(* IEC 61131-3 sources: rusty/tests/lit/single/polymorphism/interfaces, 25 files *)

(* ---- argument.st ---- *)
// RUN: %COMPILE %s && %RUN | %CHECK %s
// Scenario: Ensure interface references passed as VAR_INPUT arguments are correctly dispatched to the
// implementing function block's method.

INTERFACE IA
    METHOD foo
    END_METHOD
END_INTERFACE

INTERFACE IB
    METHOD bar
        VAR_INPUT
            refIA: IA;
        END_VAR
    END_METHOD
END_INTERFACE

FUNCTION_BLOCK FbA IMPLEMENTS IA
    METHOD foo
        printf('FbA::foo$N');
    END_METHOD
END_FUNCTION_BLOCK

FUNCTION_BLOCK FbB IMPLEMENTS IB
    VAR_INPUT
        refIA: IA;
    END_VAR

    METHOD bar
        VAR_INPUT
            refIA: IA;
        END_VAR

        refIA.foo();
        printf('FbB::bar$N');
    END_METHOD

    refIA.foo();
END_FUNCTION_BLOCK

FUNCTION main
    VAR
        instanceFbA: FbA;
        instanceFbB: FbB;
    END_VAR

    // CHECK: FbA::foo
    instanceFbB(refIA := instanceFbA);

    // CHECK-NEXT: FbA::foo
    // CHECK-NEXT: FbB::bar
    instanceFbB.bar(refIA := instanceFbA);
END_FUNCTION

(* ---- argument_implicit.st ---- *)
// RUN: %COMPILE %s && %RUN | %CHECK %s
// Scenario: FbA implements IA, FbB extends FbA and implicitly implements IA. Both should be passable as
// interface-typed arguments, with FbB's overridden method dispatched correctly.

INTERFACE IA
    METHOD foo
    END_METHOD
END_INTERFACE

FUNCTION_BLOCK FbA IMPLEMENTS IA
    METHOD foo
        printf('FbA::foo$N');
    END_METHOD
END_FUNCTION_BLOCK

FUNCTION_BLOCK FbB EXTENDS FbA
    METHOD foo
        printf('FbB::foo$N');
    END_METHOD
END_FUNCTION_BLOCK

FUNCTION_BLOCK FbC EXTENDS FbB
END_FUNCTION_BLOCK

FUNCTION_BLOCK FbConsumer
    METHOD bar
        VAR_INPUT
            refIA: IA;
        END_VAR

        refIA.foo();
    END_METHOD
END_FUNCTION_BLOCK

FUNCTION main
    VAR
        instanceFbA: FbA;
        instanceFbB: FbB;
        instanceFbC: FbC;
        consumer: FbConsumer;
    END_VAR

    // CHECK: FbA::foo
    consumer.bar(refIA := instanceFbA);

    // CHECK-NEXT: FbB::foo
    consumer.bar(refIA := instanceFbB);

    // FbC inherits FbB's override
    // CHECK-NEXT: FbB::foo
    consumer.bar(refIA := instanceFbC);
END_FUNCTION

(* ---- argument_mixed.st ---- *)
// RUN: %COMPILE %s && %RUN | %CHECK %s
// Scenario: A method takes a mix of interface-typed and non-interface-typed parameters. Only the
// interface-typed arguments should be wrapped in a fat pointer; the rest remain untouched.

INTERFACE IA
    METHOD foo
    END_METHOD
END_INTERFACE

FUNCTION_BLOCK FbA IMPLEMENTS IA
    METHOD foo
        printf('FbA::foo$N');
    END_METHOD
END_FUNCTION_BLOCK

FUNCTION_BLOCK FbConsumer
    METHOD bar
        VAR_INPUT
            x: DINT;
            refIA: IA;
            y: DINT;
        END_VAR

        printf('x=%d, y=%d$N', x, y);
        refIA.foo();
    END_METHOD
END_FUNCTION_BLOCK

FUNCTION main
    VAR
        instanceFbA: FbA;
        consumer: FbConsumer;
    END_VAR

    // CHECK: x=1, y=2
    // CHECK-NEXT: FbA::foo
    consumer.bar(x := 1, refIA := instanceFbA, y := 2);
END_FUNCTION

(* ---- argument_positional.st ---- *)
// RUN: %COMPILE %s && %RUN | %CHECK %s
// Scenario: Interface references passed as positional (unnamed) VAR_INPUT arguments are correctly wrapped
// in a fat pointer and dispatched to the implementing function block's method.

INTERFACE IA
    METHOD foo
    END_METHOD
END_INTERFACE

FUNCTION_BLOCK FbA IMPLEMENTS IA
    METHOD foo
        printf('FbA::foo$N');
    END_METHOD
END_FUNCTION_BLOCK

FUNCTION_BLOCK FbB IMPLEMENTS IA
    METHOD foo
        printf('FbB::foo$N');
    END_METHOD
END_FUNCTION_BLOCK

FUNCTION_BLOCK FbConsumer
    METHOD bar
        VAR_INPUT
            refIA: IA;
        END_VAR

        refIA.foo();
    END_METHOD
END_FUNCTION_BLOCK

FUNCTION main
    VAR
        instanceFbA: FbA;
        instanceFbB: FbB;
        consumer: FbConsumer;
    END_VAR

    // CHECK: FbA::foo
    consumer.bar(instanceFbA);

    // CHECK-NEXT: FbB::foo
    consumer.bar(instanceFbB);
END_FUNCTION

(* ---- argument_sequential.st ---- *)
// RUN: %COMPILE %s && %RUN | %CHECK %s
// Scenario: Multiple sequential calls pass different concrete types to the same interface-typed parameter.
// The single __tmp variable is reused across calls — each call should dispatch to the correct implementation.

INTERFACE IA
    METHOD foo
    END_METHOD
END_INTERFACE

FUNCTION_BLOCK FbA IMPLEMENTS IA
    METHOD foo
        printf('FbA::foo$N');
    END_METHOD
END_FUNCTION_BLOCK

FUNCTION_BLOCK FbB IMPLEMENTS IA
    METHOD foo
        printf('FbB::foo$N');
    END_METHOD
END_FUNCTION_BLOCK

FUNCTION_BLOCK FbC IMPLEMENTS IA
    METHOD foo
        printf('FbC::foo$N');
    END_METHOD
END_FUNCTION_BLOCK

FUNCTION_BLOCK FbConsumer
    METHOD bar
        VAR_INPUT
            refIA: IA;
        END_VAR

        refIA.foo();
    END_METHOD
END_FUNCTION_BLOCK

FUNCTION main
    VAR
        instanceFbA: FbA;
        instanceFbB: FbB;
        instanceFbC: FbC;
        consumer: FbConsumer;
    END_VAR

    // CHECK: FbA::foo
    consumer.bar(refIA := instanceFbA);

    // CHECK-NEXT: FbB::foo
    consumer.bar(refIA := instanceFbB);

    // CHECK-NEXT: FbC::foo
    consumer.bar(refIA := instanceFbC);

    // Back to FbA to confirm __tmp is correctly overwritten
    // CHECK-NEXT: FbA::foo
    consumer.bar(refIA := instanceFbA);
END_FUNCTION

(* ---- combined_aggregate_return_mixed_args.st ---- *)
// RUN: %COMPILE %s && %RUN | %CHECK %s
// Scenario: A method returns a STRUCT (aggregate) and takes a mix of scalar, interface, and multiple
// different interface-typed parameters. Tests both positional (unnamed) and named arguments with
// completely reordered parameter positions to verify that fat pointer wrapping targets the correct
// parameters regardless of call-site argument order.

TYPE Result :
    STRUCT
        summary: STRING;
        total: DINT;
    END_STRUCT
END_TYPE

INTERFACE IA
    METHOD describe : STRING
    END_METHOD
END_INTERFACE

INTERFACE IB
    METHOD value : DINT
    END_METHOD
END_INTERFACE

INTERFACE IC
    METHOD combine : Result
        VAR_INPUT
            x: DINT;
            a: IA;
            y: REAL;
            b: IB;
            label: STRING;
        END_VAR
    END_METHOD
END_INTERFACE

FUNCTION_BLOCK FbA IMPLEMENTS IA
    METHOD describe : STRING
        describe := 'FbA';
    END_METHOD
END_FUNCTION_BLOCK

FUNCTION_BLOCK FbB IMPLEMENTS IB
    METHOD value : DINT
        value := 100;
    END_METHOD
END_FUNCTION_BLOCK

FUNCTION_BLOCK FbC IMPLEMENTS IC
    METHOD combine : Result
        VAR_INPUT
            x: DINT;
            a: IA;
            y: REAL;
            b: IB;
            label: STRING;
        END_VAR

        // Dispatch through both interface arguments to verify their fat pointers are valid
        combine.summary := CONCAT(label, ': ');
        combine.summary := CONCAT(combine.summary, a.describe());
        combine.total := x + b.value() + REAL_TO_DINT(y);
    END_METHOD
END_FUNCTION_BLOCK

FUNCTION main
    VAR
        fa: FbA;
        fb: FbB;
        fc: FbC;
        ref_c: IC;
        result: Result;
    END_VAR

    ref_c := fc;

    // Positional (unnamed) arguments: x=10, a=fa, y=3.0, b=fb, label='test'
    // CHECK: test: FbA, 113
    result := ref_c.combine(10, fa, 3.0, fb, 'test');
    printf('%s, %d$N', result.summary, result.total);

    // Named arguments in completely different order from declaration
    // CHECK-NEXT: named: FbA, 125
    result := ref_c.combine(label := 'named', b := fb, y := 5.0, x := 20, a := fa);
    printf('%s, %d$N', result.summary, result.total);

    // Named arguments in yet another order, partial overlap with declaration order
    // CHECK-NEXT: mixed: FbA, 130
    result := ref_c.combine(a := fa, x := 30, label := 'mixed', y := 0.0, b := fb);
    printf('%s, %d$N', result.summary, result.total);
END_FUNCTION

(* ---- combined_function_aggregate_return_with_interface_argument.st ---- *)
// RUN: %COMPILE %s && %RUN | %CHECK %s
// Scenario: A free FUNCTION (not a method on an interface) returns an aggregate type (STRING) and takes
// an interface-typed VAR_INPUT. This tests the interaction between AggregateTypeLowerer and
// InterfaceDispatchLowerer for plain function calls where the callee is known statically but the
// argument still needs fat pointer wrapping.

INTERFACE IA
    METHOD name : STRING
    END_METHOD
END_INTERFACE

FUNCTION_BLOCK FbA IMPLEMENTS IA
    METHOD name : STRING
        name := 'FbA';
    END_METHOD
END_FUNCTION_BLOCK

FUNCTION_BLOCK FbB IMPLEMENTS IA
    METHOD name : STRING
        name := 'FbB';
    END_METHOD
END_FUNCTION_BLOCK

// Free function with aggregate return + interface parameter
FUNCTION format_greeting : STRING
    VAR_INPUT
        prefix: STRING;
        iface: IA;
        suffix: STRING;
    END_VAR

    format_greeting := CONCAT(prefix, iface.name());
    format_greeting := CONCAT(format_greeting, suffix);
END_FUNCTION

FUNCTION main
    VAR
        a: FbA;
        b: FbB;
        result: STRING;
    END_VAR

    // Positional call with concrete FbA instance
    // CHECK: [Hello FbA!]
    result := format_greeting('[Hello ', a, '!]');
    printf('%s$N', result);

    // Positional call with concrete FbB instance
    // CHECK-NEXT: [Hello FbB!]
    result := format_greeting('[Hello ', b, '!]');
    printf('%s$N', result);

    // Named call with reordered arguments
    // CHECK-NEXT: (Greetings FbA.)
    result := format_greeting(suffix := '.)', iface := a, prefix := '(Greetings ');
    printf('%s$N', result);

    // Named call with yet another order
    // CHECK-NEXT: {Hi FbB}
    result := format_greeting(iface := b, suffix := '}', prefix := '{Hi ');
    printf('%s$N', result);
END_FUNCTION

(* ---- combined_string_return_with_interface_argument.st ---- *)
// RUN: %COMPILE %s && %RUN | %CHECK %s
// Scenario: An interface method returns an aggregate type (STRING) and also takes an interface-typed
// argument. Both the aggregate return lowering and fat pointer wrapping must cooperate: the fat pointer
// preamble must execute before the call, and the aggregate alloca must also be set up before the call.
// This is the exact scenario that was broken when AggregateTypeLowerer ran in post_index, causing the
// interface argument to receive wrong type hints and skip fat pointer wrapping.

INTERFACE IA
    METHOD greet : STRING
        VAR_INPUT
            other: IA;
        END_VAR
    END_METHOD

    METHOD name : STRING
    END_METHOD
END_INTERFACE

FUNCTION_BLOCK FbA IMPLEMENTS IA
    METHOD greet : STRING
        VAR_INPUT
            other: IA;
        END_VAR
        greet := 'FbA says hello to ';
        // Dispatch through the interface argument to verify the fat pointer is valid
        greet := CONCAT(greet, other.name());
    END_METHOD

    METHOD name : STRING
        name := 'FbA';
    END_METHOD
END_FUNCTION_BLOCK

FUNCTION_BLOCK FbB IMPLEMENTS IA
    METHOD greet : STRING
        VAR_INPUT
            other: IA;
        END_VAR
        greet := 'FbB says hello to ';
        greet := CONCAT(greet, other.name());
    END_METHOD

    METHOD name : STRING
        name := 'FbB';
    END_METHOD
END_FUNCTION_BLOCK

FUNCTION main
    VAR
        a: FbA;
        b: FbB;
        ref_a: IA;
        ref_b: IA;
        result: STRING;
    END_VAR

    ref_a := a;
    ref_b := b;

    // Method returns STRING (aggregate) and takes an interface argument;
    // the argument must be wrapped in a fat pointer and dispatch through it.
    // CHECK: FbA says hello to FbB
    result := ref_a.greet(b);
    printf('%s$N', result);

    // CHECK-NEXT: FbB says hello to FbA
    result := ref_b.greet(a);
    printf('%s$N', result);

    // Pass an already-interface-typed variable as the argument
    // CHECK-NEXT: FbA says hello to FbB
    result := ref_a.greet(ref_b);
    printf('%s$N', result);
END_FUNCTION

(* ---- combined_struct_return_with_interface_argument.st ---- *)
// RUN: %COMPILE %s && %RUN | %CHECK %s
// Scenario: An interface method returns a user-defined STRUCT (aggregate) and takes an interface-typed
// argument. Combines struct return lowering with fat pointer wrapping. Also tests that two different
// concrete types dispatched through the same interface produce distinct results.

TYPE Pair :
    STRUCT
        first: STRING;
        second: STRING;
    END_STRUCT
END_TYPE

INTERFACE IA
    METHOD make_pair : Pair
        VAR_INPUT
            other: IA;
        END_VAR
    END_METHOD

    METHOD tag : STRING
    END_METHOD
END_INTERFACE

FUNCTION_BLOCK FbA IMPLEMENTS IA
    METHOD make_pair : Pair
        VAR_INPUT
            other: IA;
        END_VAR
        make_pair.first := 'FbA';
        make_pair.second := other.tag();
    END_METHOD

    METHOD tag : STRING
        tag := 'TagA';
    END_METHOD
END_FUNCTION_BLOCK

FUNCTION_BLOCK FbB IMPLEMENTS IA
    METHOD make_pair : Pair
        VAR_INPUT
            other: IA;
        END_VAR
        make_pair.first := 'FbB';
        make_pair.second := other.tag();
    END_METHOD

    METHOD tag : STRING
        tag := 'TagB';
    END_METHOD
END_FUNCTION_BLOCK

FUNCTION main
    VAR
        a: FbA;
        b: FbB;
        ref_a: IA;
        ref_b: IA;
        result: Pair;
    END_VAR

    ref_a := a;
    ref_b := b;

    // FbA.make_pair dispatches other.tag() through FbB's vtable
    // CHECK: first=FbA, second=TagB
    result := ref_a.make_pair(b);
    printf('first=%s, second=%s$N', result.first, result.second);

    // FbB.make_pair dispatches other.tag() through FbA's vtable
    // CHECK-NEXT: first=FbB, second=TagA
    result := ref_b.make_pair(a);
    printf('first=%s, second=%s$N', result.first, result.second);

    // Named argument
    // CHECK-NEXT: first=FbA, second=TagA
    result := ref_a.make_pair(other := a);
    printf('first=%s, second=%s$N', result.first, result.second);
END_FUNCTION

(* ---- conversion_of_base_typed_instance.st ---- *)
// RUN: %COMPILE %s && %RUN | %CHECK %s
// Scenario: An instance whose declared type is a base (`THIS^`, `ptr^`, a `REFERENCE TO`) is converted to an
// interface, by assignment or as an argument. The fat pointer must carry the itable of the actual instance,
// so a derived override runs. This also holds for interfaces added at a derived level, for an upcast to a
// parent interface after the conversion, and for classes. A plain instance keeps the itable of its type.

INTERFACE ISpeaker
    METHOD say : DINT
    END_METHOD
END_INTERFACE

INTERFACE ILoud EXTENDS ISpeaker
    METHOD shout : DINT
    END_METHOD
END_INTERFACE

INTERFACE ITagged
    METHOD tag : DINT
    END_METHOD
END_INTERFACE

FUNCTION speak : DINT
    VAR_INPUT
        s : ISpeaker;
    END_VAR

    speak := s.say();
END_FUNCTION

FUNCTION_BLOCK Dog IMPLEMENTS ILoud
    METHOD say : DINT
        say := 1;
    END_METHOD

    METHOD shout : DINT
        shout := 10;
    END_METHOD

    METHOD viaAssignment : DINT
        VAR
            s : ISpeaker;
        END_VAR

        s := THIS^;
        viaAssignment := s.say();
    END_METHOD

    METHOD viaArgument : DINT
        viaArgument := speak(THIS^);
    END_METHOD

    METHOD viaUpcast : DINT
        VAR
            l : ILoud;
            s : ISpeaker;
        END_VAR

        l := THIS^;
        s := l;
        viaUpcast := l.shout() + s.say();
    END_METHOD
END_FUNCTION_BLOCK

FUNCTION_BLOCK Puppy EXTENDS Dog IMPLEMENTS ITagged
    METHOD say : DINT
        say := 2;
    END_METHOD

    METHOD tag : DINT
        tag := 200;
    END_METHOD

    METHOD viaDerivedInterface : DINT
        VAR
            t : ITagged;
        END_VAR

        t := THIS^;
        viaDerivedInterface := t.tag();
    END_METHOD
END_FUNCTION_BLOCK

FUNCTION_BLOCK Pup EXTENDS Puppy
    METHOD say : DINT
        say := 3;
    END_METHOD

    METHOD shout : DINT
        shout := 30;
    END_METHOD

    METHOD tag : DINT
        tag := 300;
    END_METHOD
END_FUNCTION_BLOCK

CLASS Cat IMPLEMENTS ISpeaker
    METHOD say : DINT
        say := 4;
    END_METHOD
END_CLASS

CLASS Kitten EXTENDS Cat
    METHOD say : DINT
        say := 5;
    END_METHOD
END_CLASS

FUNCTION main : DINT
    VAR
        d : Dog;
        p : Puppy;
        g : Pup;
        k : Kitten;
        s : ISpeaker;
        pd : POINTER TO Dog;
        rd : REFERENCE TO Dog;
        pc : POINTER TO Cat;
        dogs : ARRAY[1..2] OF POINTER TO Dog;
    END_VAR

    // CHECK: assignment: 1 2 3
    printf('assignment: %d %d %d$N', d.viaAssignment(), p.viaAssignment(), g.viaAssignment());

    // CHECK: argument: 1 2 3
    printf('argument: %d %d %d$N', d.viaArgument(), p.viaArgument(), g.viaArgument());

    // CHECK: upcast: 11 12 33
    printf('upcast: %d %d %d$N', d.viaUpcast(), p.viaUpcast(), g.viaUpcast());

    // CHECK: derived interface: 200 300
    printf('derived interface: %d %d$N', p.viaDerivedInterface(), g.viaDerivedInterface());

    // CHECK: pointer: 3 3
    pd := ADR(g);
    s := pd^;
    printf('pointer: %d %d$N', s.say(), speak(pd^));

    // CHECK: reference: 2 2
    rd REF= p;
    s := rd;
    printf('reference: %d %d$N', s.say(), speak(rd));

    // CHECK: array of pointers: 1 3
    dogs[1] := ADR(d);
    dogs[2] := ADR(g);
    printf('array of pointers: %d %d$N', speak(dogs[1]^), speak(dogs[2]^));

    // CHECK: class: 5
    pc := ADR(k);
    s := pc^;
    printf('class: %d$N', s.say());

    // CHECK: exact: 1 2
    s := d;
    printf('exact: %d %d$N', s.say(), speak(p));
END_FUNCTION

(* ---- dispatch_conditional.st ---- *)
// RUN: %COMPILE %s && %RUN | %CHECK %s
// Scenario: Different concrete types are assigned to an interface variable based on a runtime condition.
// The method is then called after the branch, ensuring dispatch is truly dynamic and not resolved at
// compile time.

INTERFACE IA
    METHOD identify
    END_METHOD
END_INTERFACE

FUNCTION_BLOCK FbAlpha IMPLEMENTS IA
    METHOD identify
        printf('Alpha$N');
    END_METHOD
END_FUNCTION_BLOCK

FUNCTION_BLOCK FbBravo IMPLEMENTS IA
    METHOD identify
        printf('Bravo$N');
    END_METHOD
END_FUNCTION_BLOCK

FUNCTION_BLOCK FbCharlie IMPLEMENTS IA
    METHOD identify
        printf('Charlie$N');
    END_METHOD
END_FUNCTION_BLOCK

FUNCTION pick_and_call
    VAR_INPUT
        selector: DINT;
    END_VAR

    VAR
        alpha: FbAlpha;
        bravo: FbBravo;
        charlie: FbCharlie;
        reference: IA;
    END_VAR

    IF selector = 1 THEN
        reference := alpha;
    ELSIF selector = 2 THEN
        reference := bravo;
    ELSE
        reference := charlie;
    END_IF;

    reference.identify();
END_FUNCTION

FUNCTION pick_case
    VAR_INPUT
        selector: DINT;
    END_VAR

    VAR
        alpha: FbAlpha;
        bravo: FbBravo;
        charlie: FbCharlie;
        reference: IA;
    END_VAR

    CASE selector OF
        1: reference := alpha;
        2: reference := bravo;
    ELSE
        reference := charlie;
    END_CASE;

    reference.identify();
END_FUNCTION

FUNCTION main
    // IF-based selection
    // CHECK: Alpha
    pick_and_call(1);

    // CHECK-NEXT: Bravo
    pick_and_call(2);

    // CHECK-NEXT: Charlie
    pick_and_call(3);

    // CASE-based selection
    // CHECK-NEXT: Alpha
    pick_case(1);

    // CHECK-NEXT: Bravo
    pick_case(2);

    // CHECK-NEXT: Charlie
    pick_case(99);
END_FUNCTION

(* ---- dispatch_member_variable.st ---- *)
// RUN: %COMPILE %s && %RUN | %CHECK %s
// Scenario: A function block stores an interface reference as a member variable. A concrete instance is
// assigned to it, and dispatch happens through the stored reference. The fat pointer must survive being
// written to and read back from the FB's struct fields.

INTERFACE IA
    METHOD greet
    END_METHOD
END_INTERFACE

FUNCTION_BLOCK FbHello IMPLEMENTS IA
    METHOD greet
        printf('Hello$N');
    END_METHOD
END_FUNCTION_BLOCK

FUNCTION_BLOCK FbWorld IMPLEMENTS IA
    METHOD greet
        printf('World$N');
    END_METHOD
END_FUNCTION_BLOCK

FUNCTION_BLOCK FbConsumer
    VAR
        stored: IA;
    END_VAR

    METHOD store
        VAR_INPUT
            ref: IA;
        END_VAR

        stored := ref;
    END_METHOD

    METHOD invoke
        stored.greet();
    END_METHOD
END_FUNCTION_BLOCK

FUNCTION main
    VAR
        hello: FbHello;
        world: FbWorld;
        consumer: FbConsumer;
    END_VAR

    // Store FbHello, dispatch through stored member
    // CHECK: Hello
    consumer.store(hello);
    consumer.invoke();

    // Reassign to FbWorld, dispatch again
    // CHECK-NEXT: World
    consumer.store(world);
    consumer.invoke();

    // Back to FbHello to confirm no stale pointer
    // CHECK-NEXT: Hello
    consumer.store(hello);
    consumer.invoke();
END_FUNCTION

(* ---- dispatch_recursive.st ---- *)
// RUN: %COMPILE %s && %RUN | %CHECK %s
// Scenario: An interface method implementation dispatches through another interface reference passed as an
// argument, forming a chain of virtual calls. Additionally, a countdown pattern is used where an FB calls
// back into itself through an interface reference, testing re-entrant dispatch.

INTERFACE ICounter
    METHOD countdown
        VAR_INPUT
            n: DINT;
            partner: ICounter;
        END_VAR
    END_METHOD
END_INTERFACE

// FbEven prints on even numbers and delegates the next step to its partner
FUNCTION_BLOCK FbEven IMPLEMENTS ICounter
    METHOD countdown
        VAR_INPUT
            n: DINT;
            partner: ICounter;
        END_VAR

        IF n <= 0 THEN
            printf('done$N');
            RETURN;
        END_IF;

        printf('Even::%d$N', n);
        partner.countdown(n - 1, partner);
    END_METHOD
END_FUNCTION_BLOCK

// FbOdd prints on odd numbers and delegates the next step to its partner
FUNCTION_BLOCK FbOdd IMPLEMENTS ICounter
    METHOD countdown
        VAR_INPUT
            n: DINT;
            partner: ICounter;
        END_VAR

        IF n <= 0 THEN
            printf('done$N');
            RETURN;
        END_IF;

        printf('Odd::%d$N', n);
        partner.countdown(n - 1, partner);
    END_METHOD
END_FUNCTION_BLOCK

// FbSelf always delegates back to itself through the interface, testing re-entrant dispatch
FUNCTION_BLOCK FbSelf IMPLEMENTS ICounter
    METHOD countdown
        VAR_INPUT
            n: DINT;
            partner: ICounter;
        END_VAR

        IF n <= 0 THEN
            printf('done$N');
            RETURN;
        END_IF;

        printf('Self::%d$N', n);
        partner.countdown(n - 1, partner);
    END_METHOD
END_FUNCTION_BLOCK

FUNCTION main
    VAR
        even: FbEven;
        odd: FbOdd;
        self: FbSelf;
        refEven: ICounter;
        refOdd: ICounter;
        refSelf: ICounter;
    END_VAR

    refEven := even;
    refOdd := odd;
    refSelf := self;

    // Alternating dispatch: Even starts, delegates to Odd, which delegates to itself, etc.
    // CHECK: Even::3
    // CHECK-NEXT: Odd::2
    // CHECK-NEXT: Odd::1
    // CHECK-NEXT: done
    refEven.countdown(3, refOdd);

    // Self-referential: FbSelf dispatches back into itself through the interface
    // CHECK-NEXT: Self::3
    // CHECK-NEXT: Self::2
    // CHECK-NEXT: Self::1
    // CHECK-NEXT: done
    refSelf.countdown(3, refSelf);
END_FUNCTION

(* ---- hierarchy_diamond.st ---- *)
// RUN: %COMPILE %s && %RUN | %CHECK %s
// Scenario: Classic diamond pattern inheritance hierachy between interfaces. Should assert that even with
// multi inheritance dynamic dispatch works correctly.
// A
// / \
// B C
// \ /
// DD

INTERFACE A
    METHOD foo
    END_METHOD
END_INTERFACE

INTERFACE B EXTENDS A
    METHOD bar
    END_METHOD
END_INTERFACE

INTERFACE C EXTENDS A
    METHOD baz
    END_METHOD
END_INTERFACE

INTERFACE DD EXTENDS B, C
    METHOD qux
    END_METHOD
END_INTERFACE

FUNCTION_BLOCK FbA IMPLEMENTS A
    METHOD foo
        printf('FbA::foo$N');
    END_METHOD
END_FUNCTION_BLOCK

FUNCTION_BLOCK FbB IMPLEMENTS B
    METHOD foo
        printf('FbB::foo$N');
    END_METHOD

    METHOD bar
        printf('FbB::bar$N');
    END_METHOD
END_FUNCTION_BLOCK

FUNCTION_BLOCK FbC IMPLEMENTS C
    METHOD foo
        printf('FbC::foo$N');
    END_METHOD

    METHOD baz
        printf('FbC::baz$N');
    END_METHOD
END_FUNCTION_BLOCK

FUNCTION_BLOCK FbD IMPLEMENTS DD
    METHOD foo
        printf('FbD::foo$N');
    END_METHOD

    METHOD bar
        printf('FbD::bar$N');
    END_METHOD

    METHOD baz
        printf('FbD::baz$N');
    END_METHOD

    METHOD qux
        printf('FbD::qux$N');
    END_METHOD
END_FUNCTION_BLOCK

FUNCTION main
    VAR
        refA: A;
        refB: B;
        refC: C;
        refD: DD;

        instanceA: FbA;
        instanceB: FbB;
        instanceC: FbC;
        instanceD: FbD;
    END_VAR

    // ~~ refA := instance{A,B,C,DD} ~~
    refA := instanceA;
    refA.foo(); // CHECK: FbA::foo

    refA := instanceB;
    refA.foo(); // CHECK-NEXT: FbB::foo

    refA := instanceC;
    refA.foo(); // CHECK-NEXT: FbC::foo

    refA := instanceD;
    refA.foo(); // CHECK-NEXT: FbD::foo

    // ~~ refB := instance{B,DD} ~~
    refB := instanceB;
    refB.foo(); // CHECK-NEXT: FbB::foo
    refB.bar(); // CHECK-NEXT: FbB::bar

    refB := instanceD;
    refB.foo(); // CHECK-NEXT: FbD::foo
    refB.bar(); // CHECK-NEXT: FbD::bar

    // ~~ refC := instance{C,DD} ~~
    refC := instanceC;
    refC.foo(); // CHECK-NEXT: FbC::foo
    refC.baz(); // CHECK-NEXT: FbC::baz

    refC := instanceD;
    refC.foo(); // CHECK-NEXT: FbD::foo
    refC.baz(); // CHECK-NEXT: FbD::baz

    // ~~ refD := instance{DD} ~~
    refD := instanceD;
    refD.foo(); // CHECK-NEXT: FbD::foo
    refD.bar(); // CHECK-NEXT: FbD::bar
    refD.baz(); // CHECK-NEXT: FbD::baz
    refD.qux(); // CHECK-NEXT: FbD::qux
END_FUNCTION

(* ---- hierarchy_implicit.st ---- *)
// RUN: %COMPILE %s && %RUN | %CHECK %s
// Scenario: FbA is the only POU which directly implements interface A. FbB and FbC indirectly implement the
// interface by extending from FbA. Implicitly, this means FbB and FbC can be assigned to variables of type
// interface A.

INTERFACE A
    METHOD id
    END_METHOD
END_INTERFACE

// Only FbA implements A directly
FUNCTION_BLOCK FbA IMPLEMENTS A
    METHOD uniqueA1
    END_METHOD

    METHOD id
        printf('FbA$N');
    END_METHOD
END_FUNCTION_BLOCK

// FbB implicitly implements A via FbA (overridden)
FUNCTION_BLOCK FbB EXTENDS FbA
    METHOD id
        printf('FbB$N');
    END_METHOD

    METHOD uniqueB2
    END_METHOD
END_FUNCTION_BLOCK

// FbC implicitly implements A via FbB (overridden)
FUNCTION_BLOCK FbC EXTENDS FbB
    METHOD unqiueC1
    END_METHOD

    METHOD id
        printf('FbC$N');
    END_METHOD

    METHOD unqiueC2
    END_METHOD
END_FUNCTION_BLOCK

// FbD implicitly implements A via FbC (inherited)
FUNCTION_BLOCK FbD EXTENDS FbC
END_FUNCTION_BLOCK

FUNCTION main
    VAR
        reference: A;

        instanceA: FbA;
        instanceB: FbB;
        instanceC: FbC;
        instanceD: FbD;
    END_VAR

    // CHECK: FbA
    reference := instanceA;
    reference.id();

    // CHECK-NEXT: FbB
    reference := instanceB;
    reference.id();

    // CHECK-NEXT: FbC
    reference := instanceC;
    reference.id();

    // CHECK-NEXT: FbC
    reference := instanceD;
    reference.id();
END_FUNCTION

(* ---- hierarchy_linear.st ---- *)
// RUN: %COMPILE %s && %RUN | %CHECK %s
// Scenario: (Big) linear / single inheritance hierachy between interfaces, A <- B <- C <- DD <- E <- F

INTERFACE A
    METHOD foo
    END_METHOD
END_INTERFACE

INTERFACE B EXTENDS A
    METHOD bar
    END_METHOD
END_INTERFACE

INTERFACE C EXTENDS B
    METHOD baz
    END_METHOD
END_INTERFACE

INTERFACE DD EXTENDS C
    METHOD qux
    END_METHOD
END_INTERFACE

INTERFACE E EXTENDS DD
    METHOD quux
    END_METHOD
END_INTERFACE

INTERFACE F EXTENDS E
    METHOD corge
    END_METHOD
END_INTERFACE

FUNCTION_BLOCK FbA IMPLEMENTS A
    METHOD foo
        printf('FbA::foo$N');
    END_METHOD
END_FUNCTION_BLOCK

FUNCTION_BLOCK FbB IMPLEMENTS B
    METHOD foo
        printf('FbB::foo$N');
    END_METHOD

    METHOD bar
        printf('FbB::bar$N');
    END_METHOD
END_FUNCTION_BLOCK

FUNCTION_BLOCK FbC IMPLEMENTS C
    METHOD foo
        printf('FbC::foo$N');
    END_METHOD

    METHOD bar
        printf('FbC::bar$N');
    END_METHOD

    METHOD baz
        printf('FbC::baz$N');
    END_METHOD
END_FUNCTION_BLOCK

FUNCTION_BLOCK FbD IMPLEMENTS DD
    METHOD foo
        printf('FbD::foo$N');
    END_METHOD

    METHOD bar
        printf('FbD::bar$N');
    END_METHOD

    METHOD baz
        printf('FbD::baz$N');
    END_METHOD

    METHOD qux
        printf('FbD::qux$N');
    END_METHOD
END_FUNCTION_BLOCK

FUNCTION_BLOCK FbE IMPLEMENTS E
    METHOD foo
        printf('FbE::foo$N');
    END_METHOD

    METHOD bar
        printf('FbE::bar$N');
    END_METHOD

    METHOD baz
        printf('FbE::baz$N');
    END_METHOD

    METHOD qux
        printf('FbE::qux$N');
    END_METHOD

    METHOD quux
        printf('FbE::quux$N');
    END_METHOD
END_FUNCTION_BLOCK

FUNCTION_BLOCK FbF IMPLEMENTS F
    METHOD foo
        printf('FbF::foo$N');
    END_METHOD

    METHOD bar
        printf('FbF::bar$N');
    END_METHOD

    METHOD baz
        printf('FbF::baz$N');
    END_METHOD

    METHOD qux
        printf('FbF::qux$N');
    END_METHOD

    METHOD quux
        printf('FbF::quux$N');
    END_METHOD

    METHOD corge
        printf('FbF::corge$N');
    END_METHOD
END_FUNCTION_BLOCK

FUNCTION main
    VAR
        refA: A;
        refB: B;
        refC: C;
        refD: DD;
        refE: E;
        refF: F;

        instanceA: FbA;
        instanceB: FbB;
        instanceC: FbC;
        instanceD: FbD;
        instanceE: FbE;
        instanceF: FbF;
    END_VAR

    // ~~ refA := instance{A,B,C,DD,E,F} ~~
    // CHECK: FbA::foo
    // CHECK-NEXT: FbB::foo
    // CHECK-NEXT: FbC::foo
    // CHECK-NEXT: FbD::foo
    // CHECK-NEXT: FbE::foo
    // CHECK-NEXT: FbF::foo
    refA := instanceA;
    refA.foo();

    refA := instanceB;
    refA.foo();

    refA := instanceC;
    refA.foo();

    refA := instanceD;
    refA.foo();

    refA := instanceE;
    refA.foo();

    refA := instanceF;
    refA.foo();

    // ~~ refB := instance{B,C,DD,E,F} ~~
    // CHECK-NEXT: FbB::bar
    // CHECK-NEXT: FbC::bar
    // CHECK-NEXT: FbD::bar
    // CHECK-NEXT: FbE::bar
    // CHECK-NEXT: FbF::bar
    refB := instanceB;
    refB.bar();

    refB := instanceC;
    refB.bar();

    refB := instanceD;
    refB.bar();

    refB := instanceE;
    refB.bar();

    refB := instanceF;
    refB.bar();

    // ~~ refC := instance{C,DD,E,F} ~~
    // CHECK-NEXT: FbC::baz
    // CHECK-NEXT: FbD::baz
    // CHECK-NEXT: FbE::baz
    // CHECK-NEXT: FbF::baz
    refC := instanceC;
    refC.baz();

    refC := instanceD;
    refC.baz();

    refC := instanceE;
    refC.baz();

    refC := instanceF;
    refC.baz();

    // ~~ refD := instance{DD,E,F} ~~
    // CHECK-NEXT: FbD::qux
    // CHECK-NEXT: FbE::qux
    // CHECK-NEXT: FbF::qux
    refD := instanceD;
    refD.qux();

    refD := instanceE;
    refD.qux();

    refD := instanceF;
    refD.qux();

    // ~~ refE := instance{E,F} ~~
    // CHECK-NEXT: FbE::quux
    // CHECK-NEXT: FbF::quux
    refE := instanceE;
    refE.quux();

    refE := instanceF;
    refE.quux();

    // ~~ refF := instance{F} ~~
    // CHECK-NEXT: FbF::corge
    refF := instanceF;
    refF.corge();
END_FUNCTION

(* ---- hierarchy_method_name_collision.st ---- *)
// RUN: %COMPILE %s && %RUN | %CHECK %s
// Scenario: Two unrelated interfaces define a method with the same name and signature. A single function
// block implements both. Dispatching through each interface variable should resolve to the same underlying
// method, but the vtable routing for each interface must be correct independently.

INTERFACE IA
    METHOD describe : STRING
    END_METHOD

    METHOD onlyA
    END_METHOD
END_INTERFACE

INTERFACE IB
    METHOD describe : STRING
    END_METHOD

    METHOD onlyB
    END_METHOD
END_INTERFACE

FUNCTION_BLOCK FbBoth IMPLEMENTS IA, IB
    METHOD describe : STRING
        describe := 'FbBoth::describe';
    END_METHOD

    METHOD onlyA
        printf('FbBoth::onlyA$N');
    END_METHOD

    METHOD onlyB
        printf('FbBoth::onlyB$N');
    END_METHOD
END_FUNCTION_BLOCK

FUNCTION_BLOCK FbOnlyA IMPLEMENTS IA
    METHOD describe : STRING
        describe := 'FbOnlyA::describe';
    END_METHOD

    METHOD onlyA
        printf('FbOnlyA::onlyA$N');
    END_METHOD
END_FUNCTION_BLOCK

FUNCTION_BLOCK FbOnlyB IMPLEMENTS IB
    METHOD describe : STRING
        describe := 'FbOnlyB::describe';
    END_METHOD

    METHOD onlyB
        printf('FbOnlyB::onlyB$N');
    END_METHOD
END_FUNCTION_BLOCK

FUNCTION main
    VAR
        both: FbBoth;
        onlyA: FbOnlyA;
        onlyB: FbOnlyB;

        refA: IA;
        refB: IB;
    END_VAR

    // Dispatch describe() through IA — should hit FbBoth's single implementation
    // CHECK: FbBoth::describe
    refA := both;
    printf('%s$N', refA.describe());

    // Dispatch describe() through IB — same implementation, different vtable route
    // CHECK-NEXT: FbBoth::describe
    refB := both;
    printf('%s$N', refB.describe());

    // Interface-specific methods still work
    // CHECK-NEXT: FbBoth::onlyA
    refA.onlyA();

    // CHECK-NEXT: FbBoth::onlyB
    refB.onlyB();

    // Now assign different concrete types to each interface
    // CHECK-NEXT: FbOnlyA::describe
    refA := onlyA;
    printf('%s$N', refA.describe());

    // CHECK-NEXT: FbOnlyB::describe
    refB := onlyB;
    printf('%s$N', refB.describe());

    // CHECK-NEXT: FbOnlyA::onlyA
    refA.onlyA();

    // CHECK-NEXT: FbOnlyB::onlyB
    refB.onlyB();
END_FUNCTION

(* ---- hierarchy_single.st ---- *)
// RUN: %COMPILE %s && %RUN | %CHECK %s
// Scenario: Single interface which multiple function blocks implement and as a result should all be
// assignable to the interface variable in main.

INTERFACE Identifier
    METHOD printId
    END_METHOD
END_INTERFACE

FUNCTION_BLOCK FB1 IMPLEMENTS Identifier
    METHOD printId
        printf('FB1$N');
    END_METHOD
END_FUNCTION_BLOCK

FUNCTION_BLOCK FB2 IMPLEMENTS Identifier
    METHOD printId
        printf('FB2$N');
    END_METHOD
END_FUNCTION_BLOCK

FUNCTION_BLOCK FB3 IMPLEMENTS Identifier
    METHOD printId
        printf('FB3$N');
    END_METHOD
END_FUNCTION_BLOCK

FUNCTION main
    VAR
        instanceFb1: FB1;
        instanceFb2: FB2;
        instanceFb3: FB3;

        reference: Identifier;
    END_VAR

    // CHECK: FB1
    reference := instanceFb1;
    reference.printId();

    // CHECK-NEXT: FB2
    reference := instanceFb2;
    reference.printId();

    // CHECK-NEXT: FB3
    reference := instanceFb3;
    reference.printId();
END_FUNCTION

(* ---- type_array_arguments.st ---- *)
// RUN: %COMPILE %s && %RUN | %CHECK %s
// Scenario: Ensure ARRAY[1..5] OF DINT arguments are passed correctly through interface dispatch for
// VAR_INPUT, VAR_OUTPUT, VAR_IN_OUT and mixed signatures.

TYPE DintArray5: ARRAY[1..5] OF DINT; END_TYPE

INTERFACE A
    METHOD input
        VAR_INPUT
            in: DintArray5;
        END_VAR
    END_METHOD

    METHOD output
        VAR_OUTPUT
            out: DintArray5;
        END_VAR
    END_METHOD

    METHOD inout
        VAR_IN_OUT
            inout: DintArray5;
        END_VAR
    END_METHOD

    METHOD in_out_and_inout
        VAR_INPUT
            in: DintArray5;
        END_VAR

        VAR_OUTPUT
            out: DintArray5;
        END_VAR

        VAR_IN_OUT
            inout: DintArray5;
        END_VAR
    END_METHOD
END_INTERFACE

FUNCTION_BLOCK FbA IMPLEMENTS A
    METHOD input
        VAR_INPUT
            in: DintArray5;
        END_VAR

        printf('FbA::input, in = [%d, %d, %d, %d, %d]$N',
            in[1],
            in[2],
            in[3],
            in[4],
            in[5]
        );
    END_METHOD

    METHOD output
        VAR_OUTPUT
            out: DintArray5;
        END_VAR

        printf('FbA::output, out = [%d, %d, %d, %d, %d]$N',
            out[1],
            out[2],
            out[3],
            out[4],
            out[5]
        );

        out[1] := 90;
        out[2] := 91;
        out[3] := 92;
        out[4] := 93;
        out[5] := 94;
    END_METHOD

    METHOD inout
        VAR_IN_OUT
            inout: DintArray5;
        END_VAR

        printf('FbA::inout, inout = [%d, %d, %d, %d, %d]$N',
            inout[1],
            inout[2],
            inout[3],
            inout[4],
            inout[5]
        );

        inout[1] := 80;
        inout[2] := 81;
        inout[3] := 82;
        inout[4] := 83;
        inout[5] := 84;
    END_METHOD

    METHOD in_out_and_inout
        VAR_INPUT
            in: DintArray5;
        END_VAR

        VAR_OUTPUT
            out: DintArray5;
        END_VAR

        VAR_IN_OUT
            inout: DintArray5;
        END_VAR

        printf('FbA::in_out_and_inout, in = [%d, %d, %d, %d, %d]$N',
            in[1],
            in[2],
            in[3],
            in[4],
            in[5]
        );
        printf('FbA::in_out_and_inout, out = [%d, %d, %d, %d, %d]$N',
            out[1],
            out[2],
            out[3],
            out[4],
            out[5]
        );
        printf('FbA::in_out_and_inout, inout = [%d, %d, %d, %d, %d]$N',
            inout[1],
            inout[2],
            inout[3],
            inout[4],
            inout[5]
        );

        out[1] := 70;
        out[2] := 71;
        out[3] := 72;
        out[4] := 73;
        out[5] := 74;

        inout[1] := 60;
        inout[2] := 61;
        inout[3] := 62;
        inout[4] := 63;
        inout[5] := 64;
    END_METHOD
END_FUNCTION_BLOCK

FUNCTION main
    VAR
        instance: FbA;
        reference: A;

        localInputArray: DintArray5 := [21, 22, 23, 24, 25];

        localOutputArrayClean: DintArray5 := [31, 32, 33, 34, 35];
        localOutputArray: DintArray5 := [31, 32, 33, 34, 35];

        localInOutArrayClean: DintArray5 := [41, 42, 43, 44, 45];
        localInOutArray: DintArray5 := [41, 42, 43, 44, 45];
    END_VAR

    reference := instance;

    // CHECK: FbA::input, in = [21, 22, 23, 24, 25]
    reference.input(localInputArray);

    // CHECK-NEXT: FbA::output, out = [0, 0, 0, 0, 0]
    // CHECK-NEXT: main::output = [90, 91, 92, 93, 94]
    // CHECK-NEXT: main::output = [31, 32, 33, 34, 35]
    reference.output(localOutputArray);
    printf('main::output = [%d, %d, %d, %d, %d]$N',
        localOutputArray[1],
        localOutputArray[2],
        localOutputArray[3],
        localOutputArray[4],
        localOutputArray[5]
    );
    localOutputArray := localOutputArrayClean;
    printf('main::output = [%d, %d, %d, %d, %d]$N',
        localOutputArray[1],
        localOutputArray[2],
        localOutputArray[3],
        localOutputArray[4],
        localOutputArray[5]
    );

    // CHECK-NEXT: FbA::inout, inout = [41, 42, 43, 44, 45]
    // CHECK-NEXT: main::inout = [80, 81, 82, 83, 84]
    // CHECK-NEXT: main::inout = [41, 42, 43, 44, 45]
    reference.inout(localInOutArray);
    printf('main::inout = [%d, %d, %d, %d, %d]$N',
        localInOutArray[1],
        localInOutArray[2],
        localInOutArray[3],
        localInOutArray[4],
        localInOutArray[5]
    );
    localInOutArray := localInOutArrayClean;
    printf('main::inout = [%d, %d, %d, %d, %d]$N',
        localInOutArray[1],
        localInOutArray[2],
        localInOutArray[3],
        localInOutArray[4],
        localInOutArray[5]
    );

    // CHECK-NEXT: FbA::in_out_and_inout, in = [21, 22, 23, 24, 25]
    // CHECK-NEXT: FbA::in_out_and_inout, out = [0, 0, 0, 0, 0]
    // CHECK-NEXT: FbA::in_out_and_inout, inout = [41, 42, 43, 44, 45]
    // CHECK-NEXT: main::out_after_mix = [70, 71, 72, 73, 74]
    // CHECK-NEXT: main::inout_after_mix = [60, 61, 62, 63, 64]
    reference.in_out_and_inout(localInputArray, localOutputArray, localInOutArray);
    printf('main::out_after_mix = [%d, %d, %d, %d, %d]$N',
        localOutputArray[1],
        localOutputArray[2],
        localOutputArray[3],
        localOutputArray[4],
        localOutputArray[5]
    );
    printf('main::inout_after_mix = [%d, %d, %d, %d, %d]$N',
        localInOutArray[1],
        localInOutArray[2],
        localInOutArray[3],
        localInOutArray[4],
        localInOutArray[5]
    );
END_FUNCTION

(* ---- type_array_of_interfaces.st ---- *)
// RUN: %COMPILE %s && %RUN | %CHECK %s
// Scenario: An interface hierarchy (IA <- IB <- IC) with function blocks implementing each level.
// An array of the root interface IA is populated with all concrete types — direct and indirect
// implementors — and dispatched through, testing that fat pointers in array slots handle inheritance
// correctly.

INTERFACE IA
    METHOD id : DINT
    END_METHOD
END_INTERFACE

INTERFACE IB EXTENDS IA
    METHOD label : STRING
    END_METHOD
END_INTERFACE

INTERFACE IC EXTENDS IB
    METHOD depth : DINT
    END_METHOD
END_INTERFACE

FUNCTION_BLOCK Fb1 IMPLEMENTS IA
    METHOD id : DINT
        id := 1;
    END_METHOD
END_FUNCTION_BLOCK

FUNCTION_BLOCK Fb2 IMPLEMENTS IB
    METHOD id : DINT
        id := 2;
    END_METHOD

    METHOD label : STRING
        label := 'Fb2';
    END_METHOD
END_FUNCTION_BLOCK

FUNCTION_BLOCK Fb3 IMPLEMENTS IC
    METHOD id : DINT
        id := 3;
    END_METHOD

    METHOD label : STRING
        label := 'Fb3';
    END_METHOD

    METHOD depth : DINT
        depth := 3;
    END_METHOD
END_FUNCTION_BLOCK

FUNCTION main
    VAR
        inst1: Fb1;
        inst2: Fb2;
        inst3: Fb3;

        arrA: ARRAY[1..5] OF IA;
        arrB: ARRAY[1..2] OF IB;
        i: DINT;
    END_VAR

    // All three FBs are assignable to IA (direct or indirect implementation)
    arrA[1] := inst1;
    arrA[2] := inst2;
    arrA[3] := inst3;
    arrA[4] := inst2;
    arrA[5] := inst1;

    // Iterate root interface array — each element dispatches id() correctly
    // CHECK: id=1
    // CHECK-NEXT: id=2
    // CHECK-NEXT: id=3
    // CHECK-NEXT: id=2
    // CHECK-NEXT: id=1
    FOR i := 1 TO 5 DO
        printf('id=%d$N', arrA[i].id());
    END_FOR;

    // Fb2 and Fb3 are assignable to IB (direct or indirect)
    arrB[1] := inst2;
    arrB[2] := inst3;

    // Dispatch through IB array — both id() and label() work
    // CHECK-NEXT: id=2, label=Fb2
    // CHECK-NEXT: id=3, label=Fb3
    FOR i := 1 TO 2 DO
        printf('id=%d, label=%s$N', arrB[i].id(), arrB[i].label());
    END_FOR;

    // Overwrite root array element and verify dispatch changes
    // CHECK-NEXT: id=3
    arrA[1] := inst3;
    printf('id=%d$N', arrA[1].id());
END_FUNCTION

(* ---- type_array_returns.st ---- *)
// RUN: %COMPILE %s && %RUN | %CHECK %s
// Scenario: Ensure ARRAY[1..5] OF DINT return values are passed correctly through interface dispatch.

TYPE DintArray5: ARRAY[1..5] OF DINT; END_TYPE

INTERFACE A
    METHOD return_array: DintArray5
    END_METHOD
END_INTERFACE

FUNCTION_BLOCK FbA IMPLEMENTS A
    VAR
        callCounter: DINT;
    END_VAR

    METHOD return_array: DintArray5
        callCounter := callCounter + 1;

        return_array[1] := callCounter * 10 + 1;
        return_array[2] := callCounter * 10 + 2;
        return_array[3] := callCounter * 10 + 3;
        return_array[4] := callCounter * 10 + 4;
        return_array[5] := callCounter * 10 + 5;
    END_METHOD
END_FUNCTION_BLOCK

FUNCTION main
    VAR
        instance: FbA;
        reference: A;
        result: DintArray5;
    END_VAR

    reference := instance;

    // CHECK: main::result_first = [11, 12, 13, 14, 15]
    result := reference.return_array();
    printf('main::result_first = [%d, %d, %d, %d, %d]$N',
        result[1],
        result[2],
        result[3],
        result[4],
        result[5]
    );

    // CHECK-NEXT: main::result_second = [21, 22, 23, 24, 25]
    result := reference.return_array();
    printf('main::result_second = [%d, %d, %d, %d, %d]$N',
        result[1],
        result[2],
        result[3],
        result[4],
        result[5]
    );
END_FUNCTION

(* ---- type_string_arguments.st ---- *)
// RUN: %COMPILE %s && %RUN | %CHECK %s
// Scenario: Ensure STRING arguments are passed correctly through interface dispatch for
// VAR_INPUT, VAR_OUTPUT, VAR_IN_OUT and mixed signatures.

INTERFACE A
    METHOD input
        VAR_INPUT
            in_literal: STRING;
            in_variable: STRING;
        END_VAR
    END_METHOD

    METHOD output
        VAR_OUTPUT
            out: STRING;
        END_VAR
    END_METHOD

    METHOD inout
        VAR_IN_OUT
            inout: STRING;
        END_VAR
    END_METHOD

    METHOD in_out_and_inout
        VAR_INPUT
            in_literal: STRING;
            in_variable: STRING;
        END_VAR

        VAR_OUTPUT
            out: STRING;
        END_VAR

        VAR_IN_OUT
            inout: STRING;
        END_VAR
    END_METHOD
END_INTERFACE

FUNCTION_BLOCK FbA IMPLEMENTS A
    METHOD input
        VAR_INPUT
            in_literal: STRING;
            in_variable: STRING;
        END_VAR

        printf('FbA::input, in_literal = %s$N', in_literal);
        printf('FbA::input, in_variable = %s$N', in_variable);
    END_METHOD

    METHOD output
        VAR_OUTPUT
            out: STRING;
        END_VAR

        printf('FbA::output, out = %s$N', out);
        out := 'FbA::output, dirty';
    END_METHOD

    METHOD inout
        VAR_IN_OUT
            inout: STRING;
        END_VAR

        printf('FbA::inout, inout = %s$N', inout);
        inout := 'FbA::inout, dirty';
    END_METHOD

    METHOD in_out_and_inout
        VAR_INPUT
            in_literal: STRING;
            in_variable: STRING;
        END_VAR

        VAR_OUTPUT
            out: STRING;
        END_VAR

        VAR_IN_OUT
            inout: STRING;
        END_VAR

        printf('FbA::in_out_and_inout, in_literal = %s$N', in_literal);
        printf('FbA::in_out_and_inout, in_variable = %s$N', in_variable);
        printf('FbA::in_out_and_inout, out = %s$N', out);
        printf('FbA::in_out_and_inout, inout = %s$N', inout);

        out := 'FbA::in_out_and_inout, out dirty';
        inout := 'FbA::in_out_and_inout, inout dirty';
    END_METHOD
END_FUNCTION_BLOCK

FUNCTION main
    VAR
        instance: FbA;
        reference: A;

        localInputVariable: STRING := 'main, clean';
        localOutputVariable: STRING := 'main, clean';
        localInOutVariable: STRING := 'main, clean';
    END_VAR

    reference := instance;

    // CHECK: FbA::input, in_literal = input, literal
    // CHECK-NEXT: FbA::input, in_variable = main, clean
    reference.input('input, literal', localInputVariable);

    // CHECK-NEXT: FbA::output, out =
    // CHECK-NEXT: FbA::output, dirty
    // CHECK-NEXT: main, clean
    reference.output(localOutputVariable);
    printf('%s$N', localOutputVariable);
    localOutputVariable := 'main, clean';
    printf('%s$N', localOutputVariable);

    // CHECK-NEXT: FbA::inout, inout = main, clean
    // CHECK-NEXT: FbA::inout, dirty
    // CHECK-NEXT: main, clean
    reference.inout(localInOutVariable);
    printf('%s$N', localInOutVariable);
    localInOutVariable := 'main, clean';
    printf('%s$N', localInOutVariable);

    // CHECK-NEXT: FbA::in_out_and_inout, in_literal = in_out_and_inout, literal
    // CHECK-NEXT: FbA::in_out_and_inout, in_variable = main, clean
    // CHECK-NEXT: FbA::in_out_and_inout, out =
    // CHECK-NEXT: FbA::in_out_and_inout, inout = main, clean
    // CHECK-NEXT: out = FbA::in_out_and_inout, out dirty
    // CHECK-NEXT: inout = FbA::in_out_and_inout, inout dirty
    reference.in_out_and_inout('in_out_and_inout, literal', localInputVariable, localOutputVariable, localInOutVariable);
    printf('out = %s$N', localOutputVariable);
    printf('inout = %s$N', localInOutVariable);
END_FUNCTION

(* ---- type_string_returns.st ---- *)
// RUN: %COMPILE %s && %RUN | %CHECK %s
// Scenario: Ensure STRING return values are passed correctly through interface dispatch.

INTERFACE A
    METHOD return_string: STRING
    END_METHOD
END_INTERFACE

FUNCTION_BLOCK FbA IMPLEMENTS A
    VAR
        callCounter: DINT;
    END_VAR

    METHOD return_string: STRING
        callCounter := callCounter + 1;

        IF callCounter = 1 THEN
            return_string := 'FbA::return_string, first';
        ELSE
            return_string := 'FbA::return_string, second';
        END_IF
    END_METHOD
END_FUNCTION_BLOCK

FUNCTION main
    VAR
        instance: FbA;
        reference: A;
        result: STRING;
    END_VAR

    reference := instance;

    // CHECK: main::result_first = FbA::return_string, first
    result := reference.return_string();
    printf('main::result_first = %s$N', result);

    // CHECK-NEXT: main::result_second = FbA::return_string, second
    result := reference.return_string();
    printf('main::result_second = %s$N', result);
END_FUNCTION

(* ---- type_struct_arguments.st ---- *)
// RUN: %COMPILE %s && %RUN | %CHECK %s
// Scenario: Ensure user-defined STRUCT arguments are passed correctly through interface dispatch for
// VAR_INPUT, VAR_OUTPUT, VAR_IN_OUT and mixed signatures.

TYPE User :
    STRUCT
        id: ULINT;
        name: STRING;
        fingerprint: ARRAY[1..5] OF DINT;
    END_STRUCT
END_TYPE

INTERFACE A
    METHOD input
        VAR_INPUT
            in: User;
        END_VAR
    END_METHOD

    METHOD output
        VAR_OUTPUT
            out: User;
        END_VAR
    END_METHOD

    METHOD inout
        VAR_IN_OUT
            inout: User;
        END_VAR
    END_METHOD

    METHOD in_out_and_inout
        VAR_INPUT
            in: User;
        END_VAR

        VAR_OUTPUT
            out: User;
        END_VAR

        VAR_IN_OUT
            inout: User;
        END_VAR
    END_METHOD
END_INTERFACE

FUNCTION_BLOCK FbA IMPLEMENTS A
    METHOD input
        VAR_INPUT
            in: User;
        END_VAR

        printf('FbA::input, in = (id=%d, name=%s, fp=[%d, %d, %d, %d, %d])$N',
            in.id,
            in.name,
            in.fingerprint[1],
            in.fingerprint[2],
            in.fingerprint[3],
            in.fingerprint[4],
            in.fingerprint[5]
        );
    END_METHOD

    METHOD output
        VAR_OUTPUT
            out: User;
        END_VAR

        printf('FbA::output, out = (id=%d, name=%s, fp=[%d, %d, %d, %d, %d])$N',
            out.id,
            out.name,
            out.fingerprint[1],
            out.fingerprint[2],
            out.fingerprint[3],
            out.fingerprint[4],
            out.fingerprint[5]
        );

        out.id := 900;
        out.name := 'output_dirty';
        out.fingerprint[1] := 901;
        out.fingerprint[2] := 902;
        out.fingerprint[3] := 903;
        out.fingerprint[4] := 904;
        out.fingerprint[5] := 905;
    END_METHOD

    METHOD inout
        VAR_IN_OUT
            inout: User;
        END_VAR

        printf('FbA::inout, inout = (id=%d, name=%s, fp=[%d, %d, %d, %d, %d])$N',
            inout.id,
            inout.name,
            inout.fingerprint[1],
            inout.fingerprint[2],
            inout.fingerprint[3],
            inout.fingerprint[4],
            inout.fingerprint[5]
        );

        inout.id := 800;
        inout.name := 'inout_dirty';
        inout.fingerprint[1] := 801;
        inout.fingerprint[2] := 802;
        inout.fingerprint[3] := 803;
        inout.fingerprint[4] := 804;
        inout.fingerprint[5] := 805;
    END_METHOD

    METHOD in_out_and_inout
        VAR_INPUT
            in: User;
        END_VAR

        VAR_OUTPUT
            out: User;
        END_VAR

        VAR_IN_OUT
            inout: User;
        END_VAR

        printf('FbA::in_out_and_inout, in = (id=%d, name=%s, fp=[%d, %d, %d, %d, %d])$N',
            in.id,
            in.name,
            in.fingerprint[1],
            in.fingerprint[2],
            in.fingerprint[3],
            in.fingerprint[4],
            in.fingerprint[5]
        );
        printf('FbA::in_out_and_inout, out = (id=%d, name=%s, fp=[%d, %d, %d, %d, %d])$N',
            out.id,
            out.name,
            out.fingerprint[1],
            out.fingerprint[2],
            out.fingerprint[3],
            out.fingerprint[4],
            out.fingerprint[5]
        );
        printf('FbA::in_out_and_inout, inout = (id=%d, name=%s, fp=[%d, %d, %d, %d, %d])$N',
            inout.id,
            inout.name,
            inout.fingerprint[1],
            inout.fingerprint[2],
            inout.fingerprint[3],
            inout.fingerprint[4],
            inout.fingerprint[5]
        );

        out.id := 700;
        out.name := 'out_dirty';
        out.fingerprint[1] := 701;
        out.fingerprint[2] := 702;
        out.fingerprint[3] := 703;
        out.fingerprint[4] := 704;
        out.fingerprint[5] := 705;

        inout.id := 600;
        inout.name := 'inout_dirty_2';
        inout.fingerprint[1] := 601;
        inout.fingerprint[2] := 602;
        inout.fingerprint[3] := 603;
        inout.fingerprint[4] := 604;
        inout.fingerprint[5] := 605;
    END_METHOD
END_FUNCTION_BLOCK

FUNCTION main
    VAR
        instance: FbA;
        reference: A;

        localInputUser: User := (id := 201, name := 'input', fingerprint := [201, 202, 203, 204, 205]);

        localOutputUserClean: User := (id := 301, name := 'output_clean', fingerprint := [301, 302, 303, 304, 305]);
        localOutputUser: User := (id := 301, name := 'output_clean', fingerprint := [301, 302, 303, 304, 305]);

        localInOutUserClean: User := (id := 401, name := 'inout_clean', fingerprint := [401, 402, 403, 404, 405]);
        localInOutUser: User := (id := 401, name := 'inout_clean', fingerprint := [401, 402, 403, 404, 405]);
    END_VAR

    reference := instance;

    // CHECK: FbA::input, in = (id=201, name=input, fp=[201, 202, 203, 204, 205])
    reference.input(localInputUser);

    // CHECK-NEXT: FbA::output, out = (id=0, name=, fp=[0, 0, 0, 0, 0])
    // CHECK-NEXT: main::output = (id=900, name=output_dirty, fp=[901, 902, 903, 904, 905])
    // CHECK-NEXT: main::output = (id=301, name=output_clean, fp=[301, 302, 303, 304, 305])
    reference.output(localOutputUser);
    printf('main::output = (id=%d, name=%s, fp=[%d, %d, %d, %d, %d])$N',
        localOutputUser.id,
        localOutputUser.name,
        localOutputUser.fingerprint[1],
        localOutputUser.fingerprint[2],
        localOutputUser.fingerprint[3],
        localOutputUser.fingerprint[4],
        localOutputUser.fingerprint[5]
    );
    localOutputUser := localOutputUserClean;
    printf('main::output = (id=%d, name=%s, fp=[%d, %d, %d, %d, %d])$N',
        localOutputUser.id,
        localOutputUser.name,
        localOutputUser.fingerprint[1],
        localOutputUser.fingerprint[2],
        localOutputUser.fingerprint[3],
        localOutputUser.fingerprint[4],
        localOutputUser.fingerprint[5]
    );

    // CHECK-NEXT: FbA::inout, inout = (id=401, name=inout_clean, fp=[401, 402, 403, 404, 405])
    // CHECK-NEXT: main::inout = (id=800, name=inout_dirty, fp=[801, 802, 803, 804, 805])
    // CHECK-NEXT: main::inout = (id=401, name=inout_clean, fp=[401, 402, 403, 404, 405])
    reference.inout(localInOutUser);
    printf('main::inout = (id=%d, name=%s, fp=[%d, %d, %d, %d, %d])$N',
        localInOutUser.id,
        localInOutUser.name,
        localInOutUser.fingerprint[1],
        localInOutUser.fingerprint[2],
        localInOutUser.fingerprint[3],
        localInOutUser.fingerprint[4],
        localInOutUser.fingerprint[5]
    );
    localInOutUser := localInOutUserClean;
    printf('main::inout = (id=%d, name=%s, fp=[%d, %d, %d, %d, %d])$N',
        localInOutUser.id,
        localInOutUser.name,
        localInOutUser.fingerprint[1],
        localInOutUser.fingerprint[2],
        localInOutUser.fingerprint[3],
        localInOutUser.fingerprint[4],
        localInOutUser.fingerprint[5]
    );

    // CHECK-NEXT: FbA::in_out_and_inout, in = (id=201, name=input, fp=[201, 202, 203, 204, 205])
    // CHECK-NEXT: FbA::in_out_and_inout, out = (id=0, name=, fp=[0, 0, 0, 0, 0])
    // CHECK-NEXT: FbA::in_out_and_inout, inout = (id=401, name=inout_clean, fp=[401, 402, 403, 404, 405])
    // CHECK-NEXT: main::out_after_mix = (id=700, name=out_dirty, fp=[701, 702, 703, 704, 705])
    // CHECK-NEXT: main::inout_after_mix = (id=600, name=inout_dirty_2, fp=[601, 602, 603, 604, 605])
    reference.in_out_and_inout(localInputUser, localOutputUser, localInOutUser);
    printf('main::out_after_mix = (id=%d, name=%s, fp=[%d, %d, %d, %d, %d])$N',
        localOutputUser.id,
        localOutputUser.name,
        localOutputUser.fingerprint[1],
        localOutputUser.fingerprint[2],
        localOutputUser.fingerprint[3],
        localOutputUser.fingerprint[4],
        localOutputUser.fingerprint[5]
    );
    printf('main::inout_after_mix = (id=%d, name=%s, fp=[%d, %d, %d, %d, %d])$N',
        localInOutUser.id,
        localInOutUser.name,
        localInOutUser.fingerprint[1],
        localInOutUser.fingerprint[2],
        localInOutUser.fingerprint[3],
        localInOutUser.fingerprint[4],
        localInOutUser.fingerprint[5]
    );
END_FUNCTION

(* ---- type_struct_returns.st ---- *)
// RUN: %COMPILE %s && %RUN | %CHECK %s
// Scenario: Ensure user-defined STRUCT return values are passed correctly through interface dispatch.

TYPE User :
    STRUCT
        id: ULINT;
        name: STRING;
        fingerprint: ARRAY[1..5] OF DINT;
    END_STRUCT
END_TYPE

INTERFACE A
    METHOD return_user: User
    END_METHOD
END_INTERFACE

FUNCTION_BLOCK FbA IMPLEMENTS A
    VAR
        callCounter: DINT;
    END_VAR

    METHOD return_user: User
        callCounter := callCounter + 1;

        IF callCounter = 1 THEN
            return_user.id := 101;
            return_user.name := 'first';
            return_user.fingerprint[1] := 101;
            return_user.fingerprint[2] := 102;
            return_user.fingerprint[3] := 103;
            return_user.fingerprint[4] := 104;
            return_user.fingerprint[5] := 105;
        ELSE
            return_user.id := 201;
            return_user.name := 'second';
            return_user.fingerprint[1] := 201;
            return_user.fingerprint[2] := 202;
            return_user.fingerprint[3] := 203;
            return_user.fingerprint[4] := 204;
            return_user.fingerprint[5] := 205;
        END_IF
    END_METHOD
END_FUNCTION_BLOCK

FUNCTION main
    VAR
        instance: FbA;
        reference: A;
        result: User;
    END_VAR

    reference := instance;

    // CHECK: main::result_first = (id=101, name=first, fp=[101, 102, 103, 104, 105])
    result := reference.return_user();
    printf('main::result_first = (id=%d, name=%s, fp=[%d, %d, %d, %d, %d])$N',
        result.id,
        result.name,
        result.fingerprint[1],
        result.fingerprint[2],
        result.fingerprint[3],
        result.fingerprint[4],
        result.fingerprint[5]
    );

    // CHECK-NEXT: main::result_second = (id=201, name=second, fp=[201, 202, 203, 204, 205])
    result := reference.return_user();
    printf('main::result_second = (id=%d, name=%s, fp=[%d, %d, %d, %d, %d])$N',
        result.id,
        result.name,
        result.fingerprint[1],
        result.fingerprint[2],
        result.fingerprint[3],
        result.fingerprint[4],
        result.fingerprint[5]
    );
END_FUNCTION
